PROGRAM main
VAR
	test_read AT %QW0 : int;
	test_coil AT %QX0.0 : bool;
END_VAR

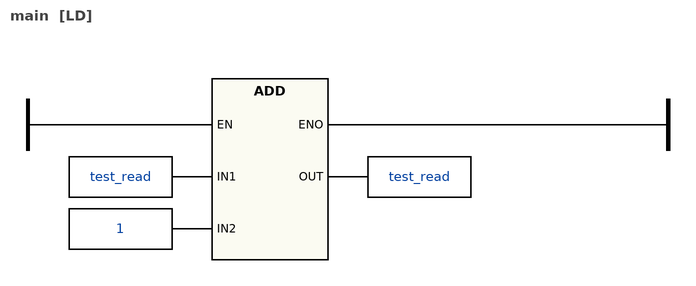
(* LD diagram, written out as Structured Text *)
test_read := test_read + 1;
END_PROGRAM
